// Generated by voz_llm_plc_agent
// Target: Siemens TIA Portal V18 - SCL external source
// Review and compile before any download to physical hardware.

FUNCTION_BLOCK "PLC_PRG"
{ S7_Optimized_Access := 'TRUE' }
VERSION : 0.1
VAR_INPUT
   I_Mode_Manual : Bool := FALSE;
   I_Mode_Auto : Bool := FALSE;
   I_Start : Bool := FALSE;
   I_Stop : Bool := FALSE;
   I_Emergency : Bool := FALSE;
   I_Auto_Motor_Command : Bool := FALSE;
   I_Manual_Motor_Command : Bool := FALSE;
END_VAR
VAR_OUTPUT
   Q_Motor_Enable : Bool := FALSE;
END_VAR
VAR
   M_ManualMode : Bool;
   M_AutoMode : Bool;
END_VAR
BEGIN
(* Selector de modo MODE_AUTO (TRUE = Automatico, FALSE = Manual): el motor sigue la orden del *)
(* modo seleccionado; la orden del otro modo no tiene efecto. *)
#M_AutoMode := #I_Mode_Auto;
#M_ManualMode := NOT #I_Mode_Auto;
#Q_Motor_Enable := ((#M_AutoMode AND #I_Auto_Motor_Command) OR (#M_ManualMode AND #I_Manual_Motor_Command)) AND NOT #I_Emergency;
END_FUNCTION_BLOCK

DATA_BLOCK "DB_PLC_PRG"
{ S7_Optimized_Access := 'TRUE' }
VERSION : 0.1
NON_RETAIN
"PLC_PRG"
BEGIN
END_DATA_BLOCK

ORGANIZATION_BLOCK "Main"
{ S7_Optimized_Access := 'TRUE' }
VERSION : 0.1
BEGIN
   "DB_PLC_PRG"(
      I_Mode_Manual := "I_Mode_Manual",
      I_Mode_Auto := "I_Mode_Auto",
      I_Start := "I_Start",
      I_Stop := "I_Stop",
      I_Emergency := "I_Emergency",
      Q_Motor_Enable => "Q_Motor_Enable",
      I_Auto_Motor_Command := "I_Auto_Motor_Command",
      I_Manual_Motor_Command := "I_Manual_Motor_Command"
   );
END_ORGANIZATION_BLOCK
